Fanuc KAREL source: kb00161.KL

PROGRAM KB00161
%NOLOCKGROUP
%ENVIRONMENT REGOPE
VAR
P1:INTEGER;P2 : XYZWPREXT;P3:INTEGER
BEGIN
--
--
P1=1
P3=1
SET_EPOS_REG(P1,P2,P3,1)
END KB00161
